# EPICS substitutions: xrmIocApp/Db/permit_lut_32R.substitutions
file "permit_lut.template"
{
	pattern {ROW0, ADDR}
	{01, 0}
	{02, 1}
	{03, 2}
	{04, 3}
	{05, 4}
	{06, 5}
	{07, 6}
	{08, 7}
	{09, 8}
	{10, 9}
	{11,10}
	{12,11}
	{13,12}
	{14,13}
	{15,14}
	{16,15}
	{17,16}
	{18,17}
	{19,18}
	{20,19}
	{21,20}
	{22,21}
	{23,22}
	{24,23}
	{25,24}
	{26,25}
	{27,26}
	{28,27}
	{29,28}
	{30,29}
	{31,30}
	{32,31}
}
